Fanuc KAREL source: ko00098.KL

PROGRAM KO00098
%STACKSIZE=65535
%PRIORITY=65535
%NOLOCKGROUP
VAR
A : INTEGER
B : INTEGER
OUT : REAL
BEGIN
A=1
B=2
-- UNRESOLVED_PC line 10 opcodes [27 27 21 64 27 21 64 76 23] marker_code=28
END KO00098
